TYPE E_Zustand :
(
	Aus := 0,
	Bereit := 1,
	Heizen := 2,
	Warnung := 3,
	Kritisch := 4,
	Notaus := 5
);
END_TYPE

(* stored: Version 1.1.0.1, ProductVersion 3.1.4024.32
   DUT E_Zustand: Id {08D95A1B-2C3D-4849-6A5B-D6E7F8091A2B} *)
